FUNCTION_BLOCK FB_Control
VAR_INPUT
END_VAR
VAR_OUTPUT
END_VAR
VAR
END_VAR

END_FUNCTION_BLOCK

(* stored: Version 1.1.0.1
   POU FB_Control: Id {2aa00cb3-4e44-47d1-aee6-f5c5ea778fd3}, SpecialFunc None *)
